(* IEC 61131-3 sources: plcassist-cli/packages/volt-lsp-iec/test-corpus/lenze-mid/Device/Plc Logic/Application/Library Manager/L_OEEA_BaseDependency, 3.26.4.8 (Lenze), 18 files *)

(* ---- GVL_CONST_PRODUCTION_LOG.gvl ---- *)
VAR_GLOBAL
	IMAXSIZEXY_TREND : INT := 100;
END_VAR

(* ---- GVL_GLOBAL_CONSTANTS.gvl ---- *)
VAR_GLOBAL
	UIMAXLOGSIZE : UINT := 50;
	IMAXFIELDS : INT := 30;
END_VAR

(* ---- GVL_MPCONSTS.gvl ---- *)
VAR_GLOBAL
	UINOOFPARTCOUNTER : UINT := 2;
	UINOOFPRODUCTIONMODES : UINT := 20;
	UINOOFDOWNTIMECATEGORIES : UINT := 99;
END_VAR

(* ---- GVL_SSCONSTS.gvl ---- *)
VAR_GLOBAL
	UINOOFSHIFTS : UINT := 3;
	UIDAYSCHEDULE : UINT := 7;
	UISHIFTNAME : UINT := 80;
	UINOOFBREAKS : UINT := 9;
END_VAR

(* ---- VERSIONCONSTANTS.gvl ---- *)
VAR_GLOBAL
	GC_BYAMOUNTOFGENERALDATA : BYTE := 50;
	GC_BYAMOUNTDOWNTIMEERRORS : BYTE := 10;
	GC_IFILTERSAMPLES : INT := 20;
END_VAR

(* ---- BOOL_TO_SQLSTRING.fun ---- *)
FUNCTION BOOL_TO_SQLSTRING : STRING
VAR_INPUT
	XBOOLVALUE : BOOL;
END_VAR
END_FUNCTION

(* ---- CALC_UNIXTIME.fun ---- *)
FUNCTION CALC_UNIXTIME : DINT
VAR_INPUT
	DTACTUALDATETIME : DATE_AND_TIME;
END_VAR
END_FUNCTION

(* ---- CONVERTDATETIME_TO_STR.fun ---- *)
FUNCTION CONVERTDATETIME_TO_STR : STRING
VAR_INPUT
	DTTIME_VALUE : DATE_AND_TIME;
END_VAR
END_FUNCTION

(* ---- CONVERTTIME_TO_STR.fun ---- *)
FUNCTION CONVERTTIME_TO_STR : STRING
VAR_INPUT
	TTIME_VALUE : TIME;
END_VAR
END_FUNCTION

(* ---- CONVERTTOD_TO_STR.fun ---- *)
FUNCTION CONVERTTOD_TO_STR : STRING
VAR_INPUT
	TODTIME_VALUE : TIME_OF_DAY;
END_VAR
END_FUNCTION

(* ---- CUTDECIMALLREALVALUE.fun ---- *)
FUNCTION CUTDECIMALLREALVALUE : LREAL
VAR_INPUT
	LRVALUE : LREAL;
	INOOFDECIMAL : INT;
END_VAR
END_FUNCTION

(* ---- CUTDECIMALREALVALUE.fun ---- *)
FUNCTION CUTDECIMALREALVALUE : REAL
VAR_INPUT
	RVALUE : REAL;
	INOOFDECIMAL : INT;
END_VAR
END_FUNCTION

(* ---- CUTREALVALUE.fun ---- *)
FUNCTION CUTREALVALUE : REAL
VAR_INPUT
	RVALUE : REAL;
	INOOFDECIMAL : INT;
	INOOFAVERAGECOUNT : INT;
END_VAR
VAR_IN_OUT
	SCCUTAVERAGEREAL : scCutAverageReal;
END_VAR
END_FUNCTION

(* ---- STRING_TO_SQLSTRING.fun ---- *)
FUNCTION STRING_TO_SQLSTRING : STRING
VAR_INPUT
	SSTRINGVALUE : STRING;
END_VAR
END_FUNCTION

(* ---- TIMEPERIOD.fun ---- *)
FUNCTION TIMEPERIOD : TIME
VAR_INPUT
	DTSTARTTIME : TIME_OF_DAY;
	DTENDTIME : TIME_OF_DAY;
END_VAR
END_FUNCTION

(* ---- TOD_TO_SECONDS.fun ---- *)
FUNCTION TOD_TO_SECONDS : DINT
VAR_INPUT
	TODTIME : TIME_OF_DAY;
END_VAR
END_FUNCTION

(* ---- TODCONCAT_SECONDVALUE.fun ---- *)
FUNCTION TODCONCAT_SECONDVALUE : TIME_OF_DAY
VAR_INPUT
	DISECONDSVALUE : DINT;
END_VAR
END_FUNCTION

(* ---- TODSPLIT_DAYCHANGECALC.fun ---- *)
FUNCTION TODSPLIT_DAYCHANGECALC : DINT
VAR_INPUT
	TODTIMEHIGH : TIME_OF_DAY;
	TODTIMELOW : TIME_OF_DAY;
	PUIHOUR : UINT;
	PUIMINUTE : UINT;
	PUISECOND : UINT;
	PUIMILLISECOND : UINT;
END_VAR
END_FUNCTION
